FUNCTION_BLOCK FB_DriveInterface
VAR_INPUT
TorqueSetpoints : ST_JointTorque;
Config           : ST_TherapyConfig;
END_VAR
VAR_OUTPUT
END_VAR
VAR
	
	lrRatedTorque_Axis1 : LREAL := 810.425; 
    lrRatedTorque_Axis2 : LREAL := 383.934;
    lrRatedTorque_Axis3 : LREAL := 382.060;
	
	fbTorqueAxis1    : MC_TorqueControl;
    fbTorqueAxis2    : MC_TorqueControl;
    fbTorqueAxis3    : MC_TorqueControl;
	lrTorqueSetpoint_Pct : ST_JointTorque;
	
	lrEffectiveSpeedHigh  : LREAL;
    lrEffectiveSpeedLow   : LREAL;
	ErrorAxisA: BOOL;
	ErrorAxisID: UDINT;
	Execute_A : BOOL ;
	Execute_B : BOOL ;
	Execute_C : BOOL ;
	TurnOnMotors: BOOL := FALSE;
	
	
	ErrorAxisID_A: UDINT;
	ErrorAxisID_B: UDINT;
	ErrorAxisB: BOOL;
	ErrorAxisC: BOOL;
	ErrorAxisID_C: UDINT;
	torqueofaxisB: BOOL;
	BisBusy: BOOL;
	BisActive: BOOL;
	torqueofaxisA: BOOL;
	AisBusy: BOOL;
	AisActive: BOOL;
END_VAR

// 1. Clamp Positive Game Limit between 0.0 and +GlobalVelocityLimit
lrEffectiveSpeedHigh := LIMIT(
    0.0, 
    ABS(Config.GlobalVelocityLimit), // THIS Data should changed based on game currently I put equal tp g;pbalspeedlimitHigh
    ABS(Config.GlobalVelocityLimit)
);

// 2. Clamp Negative Game Limit between -GlobalVelocityLimit and 0.0
lrEffectiveSpeedLow  := LIMIT(
    -ABS(Config.GlobalVelocityLimit), // THIS Data should changed based on game currently I put equal tp g;pbalspeedlimitHigh
    -ABS(Config.GlobalVelocityLimit), 
    0.0
);



// SCALING NM to Percentage
// Motor 1 (Axis 1)
lrTorqueSetpoint_Pct.M1 := (TorqueSetpoints.M1 / lrRatedTorque_Axis1) * 100.0;

// Motor 2 (Axis 2)
lrTorqueSetpoint_Pct.M2 := (TorqueSetpoints.M2 / lrRatedTorque_Axis2) * 100.0;
// Motor 3 (Axis 3)
lrTorqueSetpoint_Pct.M3 := (TorqueSetpoints.M3 / lrRatedTorque_Axis3) * 100.0;

lrTorqueSetpoint_Pct.M1 := TorqueSetpoints.M1;
lrTorqueSetpoint_Pct.M2 := TorqueSetpoints.M2;
lrTorqueSetpoint_Pct.M3 := TorqueSetpoints.M3;


// lrTorqueSetpoint_Pct.M1 := 20.0;
// lrTorqueSetpoint_Pct.M2 := 50.0;
// lrTorqueSetpoint_Pct.M3 := -50.0;	

//lrTorqueSetpoint_Pct.M1 := TorqueSetpoints.M1;
//lrTorqueSetpoint_Pct.M2 := TorqueSetpoints.M2;
//lrTorqueSetpoint_Pct.M3 := TorqueSetpoints.M3;

Execute_A := GVL_HMI.ContinueTOWorkspaceLimits;
Execute_B := GVL_HMI.ContinueTOWorkspaceLimits;
Execute_C := GVL_HMI.ContinueTOWorkspaceLimits;


fbTorqueAxis1(
    Axis             := GVL_Axes.Axis1,
    Execute          := Execute_A,                 // Keep TRUE to stay active
    ContinuousUpdate := TRUE,                 // CRITICAL: Allows changing torque every cycle
    Torque           := lrTorqueSetpoint_Pct.M1,   // Input from Jacobian
    Relative         := FALSE,  // Absolute Torque
	TorqueRamp         :=   100.0,               
    VelocityLimitHigh:= lrEffectiveSpeedHigh,        // Safety: Prevent runaway if resistance is lost
    VelocityLimitLow := lrEffectiveSpeedLow,
	InTorque => torqueofaxisA,
	Busy=> AisBusy,
	Active => AisActive,
	Error => ErrorAxisA ,
	ErrorID => ErrorAxisID_A
);

// -----------------------------------------------------------------------------
// AXIS 2 TORQUE CONTROL
// -----------------------------------------------------------------------------
fbTorqueAxis2(
    Axis             := GVL_Axes.Axis2,
    Execute          := Execute_B,
    ContinuousUpdate := TRUE,
    Torque           := lrTorqueSetpoint_Pct.M2,
    Relative         := FALSE,
	TorqueRamp         := 100.0,
    VelocityLimitHigh:= lrEffectiveSpeedHigh,        // Safety: Prevent runaway if resistance is lost
    VelocityLimitLow := lrEffectiveSpeedLow,
	InTorque => torqueofaxisB,
	Busy=> BisBusy,
	Active => BisActive,
	
	Error => ErrorAxisB ,
	ErrorID => ErrorAxisID_B
);

// -----------------------------------------------------------------------------
// AXIS 3 TORQUE CONTROL
// -----------------------------------------------------------------------------
fbTorqueAxis3(
    Axis             := GVL_Axes.Axis3,
    Execute          := Execute_C,
    ContinuousUpdate := TRUE,
    Torque           := lrTorqueSetpoint_Pct.M3,
    Relative         := FALSE,
	TorqueRamp         :=   100.0,
    VelocityLimitHigh:= lrEffectiveSpeedHigh,        // Safety: Prevent runaway if resistance is lost
    VelocityLimitLow := lrEffectiveSpeedLow,
	Error => ErrorAxisC,
	ErrorID => ErrorAxisID_C
);

// DriveMotors := TRUE;

END_FUNCTION_BLOCK

(* stored: Version 1.1.0.1, ProductVersion 3.1.4024.15
   POU FB_DriveInterface: Id {8a220163-88d7-4c61-b531-50b23c68dc6e}, SpecialFunc None *)
